(* IEC 61131-3 sources: llm-plc-st-eval/data/definitivo/qwen2.5-coder_14b/C5/zero_shot, 2 files *)

(* ---- ejec_3.st ---- *)
1. **Error en la sección CASE estado OF:**
   - **Línea:** 20-22
   - **Explicación:** En el estado 1, se activa el temporizador `t1` y se espera que termine para pasar al estado 2. Sin embargo, no se desactiva el contactor `kY` antes de activar `kD`. Esto viola la regla de que `kY` y `kD` no deben estar activos simultáneamente.
   - **Corrección:** Desactivar `kY` antes de activar `kD` en el estado 1.

2. **Error en la sección CASE estado OF:**
   - **Línea:** 25
   - **Explicación:** En el estado 2, se desactiva `kY`, pero no se asegura que `kD` se mantenga activo después de que `t1` termine. Esto podría causar un comportamiento inesperado.
   - **Corrección:** Asegurar que `kD` se mantenga activo después de que `t1` termine.

3. **Error en la sección CASE estado OF:**
   - **Línea:** 20-22
   - **Explicación:** En el estado 1, se activa el temporizador `t1` y se espera que termine para pasar al estado 2. Sin embargo, no se respetan los 100 milisegundos de tiempo muerto antes de activar `kD`.
   - **Corrección:** Añadir un temporizador adicional para gestionar el tiempo muerto de 100 milisegundos.

4. **Error en la sección IF btnParo THEN:**
   - **Línea:** 30-32
   - **Explicación:** Al pulsar `btnParo`, se desactivan `kY` y `kD`, pero no se desactiva `kM`. Esto podría causar un comportamiento inesperado.
   - **Corrección:** Añadir la desactivación de `kM` al pulsar `btnParo`.

**Correcciones propuestas:**

```iec
FUNCTION_BLOCK FB_EstrellaTriangulo
VAR_INPUT
    btnMarcha : BOOL;
    btnParo : BOOL;
END_VAR
VAR_OUTPUT
    kM : BOOL;
    kY : BOOL;
    kD : BOOL;
END_VAR
VAR
    estado : INT;
    t1 : TON;
    t2 : TON;
    t3 : TON;  // Nuevo temporizador para el tiempo muerto
END_VAR

CASE estado OF
    0:
        IF btnMarcha THEN
            kM := TRUE;
            kY := TRUE;
            estado := 1;
        END_IF
    1:
        t1(IN := TRUE, PT := T#8S);
        IF t1.Q THEN
            kY := FALSE;  // Desactivar kY antes de activar kD
            t3(IN := TRUE, PT := T#100MS);  // Iniciar temporizador para el tiempo muerto
            estado := 2;
        END_IF
    2:
        IF t3.Q THEN  // Esperar el tiempo muerto
            kD := TRUE;
        END_IF
END_CASE

IF btnParo THEN
    kM := FALSE;  // Desactivar kM al pulsar btnParo
    kY := FALSE;
    kD := FALSE;
    estado := 0;
END_IF
END_FUNCTION_BLOCK
```

(* ---- ejec_1.st ---- *)
1. **Error en la sección CASE estado OF:**
   - **Línea:** 18-20
   - **Explicación:** En el estado 1, se activa `kD` y se pasa al estado 2, pero no se desactiva `kY` antes de activar `kD`. Esto viola la condición de que `kY` y `kD` no deben estar activos simultáneamente.
   - **Corrección:** Desactivar `kY` antes de activar `kD` en el estado 1.
     ```pascal
     1:
         t1(IN := TRUE, PT := T#8S);
         IF t1.Q THEN
             kY := FALSE;  // Agregar esta línea
             kD := TRUE;
             estado := 2;
         END_IF
     ```

2. **Error en la sección CASE estado OF:**
   - **Línea:** 22
   - **Explicación:** En el estado 2, solo se desactiva `kY`, pero no se asegura que `kD` esté activo. Esto podría causar un comportamiento inesperado si `kD` no se activa correctamente.
   - **Corrección:** Asegurarse de que `kD` esté activo en el estado 2.
     ```pascal
     2:
         kY := FALSE;
         kD := TRUE;  // Asegurarse de que kD esté activo
     ```

3. **Error en la sección IF btnParo THEN:**
   - **Línea:** 26-28
   - **Explicación:** Al pulsar `btnParo`, solo se desactivan `kY` y `kD`, pero no se desactiva `kM`. Esto podría dejar el sistema en un estado inconsistente.
   - **Corrección:** Desactivar `kM` al pulsar `btnParo`.
     ```pascal
     IF btnParo THEN
         kM := FALSE;  // Agregar esta línea
         kY := FALSE;
         kD := FALSE;
         estado := 0;
     END_IF
     ```

4. **Error en la sección CASE estado OF:**
   - **Línea:** 18-20
   - **Explicación:** En el estado 1, se activa `kD` y se pasa al estado 2, pero no se respetan los 100 milisegundos de tiempo muerto antes de activar `kD`.
   - **Corrección:** Agregar un temporizador adicional para el tiempo muerto antes de activar `kD`.
     ```pascal
     VAR
         t1 : TON;
         t2 : TON;
         t3 : TON;  // Agregar temporizador t3 para el tiempo muerto
     END_VAR

     1:
         t1(IN := TRUE, PT := T#8S);
         IF t1.Q THEN
             t3(IN := TRUE, PT := T#100MS);  // Iniciar temporizador t3
             IF t3.Q THEN
                 kY := FALSE;
                 kD := TRUE;
                 estado := 2;
             END_IF
         END_IF
     ```

5. **Error en la sección CASE estado OF:**
   - **Línea:** 22
   - **Explicación:** En el estado 2, solo se desactiva `kY`, pero no se asegura que `kD` esté activo. Esto podría causar un comportamiento inesperado si `kD` no se activa correctamente.
   - **Corrección:** Asegurarse de que `kD` esté activo en el estado 2.
     ```pascal
     2:
         kY := FALSE;
         kD := TRUE;  // Asegurarse de que kD esté activo
     ```

Con estas correcciones, el programa debería implementar correctamente el arranque estrella-triángulo, respetando todas las condiciones especificadas.
